(* IEC 61131-3 sources: model-first-plc-agent-ai/results/T3-B-08, 1 file *)

(* ---- b_code.st ---- *)
FUNCTION_BLOCK TankFillingControl
VAR_INPUT
    start : BOOL;
    stop : BOOL;
    LSH : BOOL;
    LSHH : BOOL;
    TON_Duration : TIME;
    TOF_Duration : TIME;
END_VAR
VAR_OUTPUT
    fill_valve : BOOL;
    discharge_valve : BOOL;
END_VAR
VAR
    phase : INT := 0; (* 0 = idle, 1 = filling, 2 = pause *)
    filling_active : BOOL;
    ton_q : BOOL;
    tof_q : BOOL;
    filling_timer : TON;
    pause_timer : TOF;
END_VAR

(* Both timers use the activity of the filling step. *)
filling_active := (phase = 1);

filling_timer(IN := filling_active, PT := TON_Duration);
pause_timer(IN := filling_active, PT := TOF_Duration);

ton_q := filling_timer.Q;
tof_q := pause_timer.Q;

(* Stop and level interlocks take priority over every transition. *)
IF stop OR LSH OR LSHH THEN
    phase := 0;
ELSE
    CASE phase OF
        0:
            IF start THEN
                phase := 1;
            END_IF;

        1:
            IF ton_q THEN
                phase := 2;
            END_IF;

        2:
            IF NOT tof_q THEN
                phase := 1;
            END_IF;

        ELSE
            phase := 0;
    END_CASE;
END_IF;

fill_valve := (phase = 1) AND NOT stop AND NOT LSH AND NOT LSHH;
discharge_valve := FALSE;

END_FUNCTION_BLOCK

PROGRAM Main
VAR
    StartCommand AT %IX100.0 : BOOL;
    StopCommand AT %IX100.1 : BOOL;
    LSH AT %IX100.2 : BOOL;
    LSHH AT %IX100.3 : BOOL;

    FillValve AT %QX100.0 : BOOL;
    DischargeValve AT %QX100.1 : BOOL;
END_VAR
VAR
    (* Adjustable timing parameters. *)
    TON_Duration : TIME := T#5s;
    TOF_Duration : TIME := T#5s;

    start : BOOL;
    stop : BOOL;
    fill_valve : BOOL;
    discharge_valve : BOOL;

    start_edge : R_TRIG;
    tank_control : TankFillingControl;
END_VAR

start_edge(CLK := StartCommand);
start := start_edge.Q;
stop := StopCommand;

tank_control(
    start := start,
    stop := stop,
    LSH := LSH,
    LSHH := LSHH,
    TON_Duration := TON_Duration,
    TOF_Duration := TOF_Duration
);

fill_valve := tank_control.fill_valve;
discharge_valve := tank_control.discharge_valve;

FillValve := fill_valve;
DischargeValve := discharge_valve;

END_PROGRAM
